FUNCTION_BLOCK F_NOT_BOOL (* standard boolean NOT function - Simple FB mit nativer ST-Negation (kein externes F_NOT, kein Composite-Netzwerk mehr noetig) *)
  (* Standard: 61131-3; Classification: standard boolean function; Description: Copyright (c) 2011 TU Wien ACIN, HR Agrartechnik GmbH This program and the accompanying materials are made available under the terms of the Eclipse Public License 2.0 which is available at https://www.eclipse.org/legal/epl-2.0/ SPDX-License-Identifier: EPL-2.0 *)
  (* Version 3.2, 2026-10-11, Franz Höpfinger, Meisterschulen am Ostbahnhof, Von Composite FB (FBNetwork mit NOOP + Negated-Datenverbindung) auf Simple FB umgestellt: OUT := NOT IN; direkt als ST-Algorithmus. Kein internes FB mehr, keine iec61131-3-Abhaengigkeit. *)
  (* Version 3.1, 2026-10-11, Franz Höpfinger, Meisterschulen am Ostbahnhof, Interne Umsetzung wrapt jetzt NOOP (+ Negated-Attribut auf der IN-Datenverbindung) statt iec61131::bitwiseOperators::F_NOT - damit entfaellt die letzte iec61131-3-Abhaengigkeit dieses Pakets. Instanzname F_NOT auf Negate umbenannt (Type ist jetzt NOOP, Name war sonst irrefuehrend). Organization-Attribut ergaenzt (XSD-Pflichtfeld). *)
  (* Version 3.0, 2025-04-14, Patrick Aigner, Eclipse 4diac, changed package *)
  (* Version 1.0, 2011-06-21, Monika Wenger, TU Wien ACIN, initial API and implementation and/or initial documentation *)
  PACKAGE iec61131::booleanOperators;
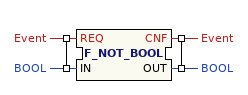
  EVENT_INPUT
    REQ WITH IN; (* Service Request *)
  END_EVENT
  EVENT_OUTPUT
    CNF WITH OUT; (* Confirmation of Requested Service *)
  END_EVENT
  VAR_INPUT
    IN : BOOL; (* Input *)
  END_VAR
  VAR_OUTPUT
    OUT : BOOL; (* Output *)
  END_VAR
  EC_STATES
    REQ : REQ -> CNF;
  END_STATES
  ALGORITHM REQ IN ST: (* Executed algorithm *)
OUT := NOT IN;
  END_ALGORITHM
END_FUNCTION_BLOCK
